Fanuc KAREL source: KT00925.KL

PROGRAM KT00925
%NOLOCKGROUP
VAR
  R1: REAL
  R2: REAL
  OUT: STRING[80]
BEGIN
  R1 = 2.0
  R2 = 3.0
  R1 = 2.0
  R2 = 3.0
  OUT = SUB_STR(R1, 1, 1)
END KT00925
